(*~
	<docu>
		<summary>
			Parameter identifiers of the "Read parameters" command (manual pp. 43-46). Every value is exchanged as LONG x1000; times in seconds, levels in the instrument units, selections as code x1000.
		</summary>
	</docu>
~*)
{attribute 'qualified_only'}
{attribute 'strict'}
TYPE eTcoAteqG6_ParameterId_v_3_5_x :
(
	None := 0,
	FillTime := 1,
	StabTime := 2,
	TestTime := 3,
	PreFillTime := 6,
	DumpTime := 9,
	CouplingTimeA := 10,
	CouplingTimeB := 11,
	PartVolume := 20,
	TestType := 21,
	InterCycleTime := 29,
	ResultHoldTime := 48,
	MinFill := 50,
	MaxFill := 51,
	PressureUnit := 53,
	TestFail := 60,
	TestRework := 61,
	RefFail := 62,
	RefRework := 63,
	SetFill := 66,
	DiffAutoResetTime := 80,
	FillMode := 103,
	ExternalDumpType := 110,
	Input7Function := 112,
	Language := 123,
	MaxPreFill := 126,
	FlowUnit := 127,
	CalibrationLeakRate := 128,
	Filter := 148,
	UnitType := 149,
	BarGraphMaxReject := 158,
	VolumeUnit := 161,
	NextProgram := 164,
	PiezoAutoZeroCycles := 165,
	PiezoAutoZeroMinutes := 166,
	DelayExt1 := 249,
	DelayExt2 := 250,
	DelayExt3 := 251,
	DelayExt4 := 252,
	DelayExt5 := 253,
	DelayExt6 := 254,
	DelayInt2 := 255,
	DelayInt1 := 256,
	DelayAux1 := 257,
	DelayAux2 := 258,
	DelayAux3 := 259,
	DelayAux4 := 260,
	TimeExt1 := 261,
	TimeExt2 := 262,
	TimeExt3 := 263,
	TimeExt4 := 264,
	TimeExt5 := 265,
	TimeExt6 := 266,
	TimeInt2 := 267,
	TimeInt1 := 268,
	TimeAux1 := 269,
	TimeAux2 := 270,
	TimeAux3 := 271,
	TimeAux4 := 272,
	PressureFilter := 274,
	CapillaryRange := 281,
	BarCodeFirstChar := 287,
	BarCodeCharCount := 288,
	BarCodeProgram := 289,
	GeneralPressureUnit := 353,
	LinePressureMin := 354,
	DisplayMode := 364,
	Input8Function := 375,
	Input9Function := 376,
	UsbMode := 379,
	SaveOn := 412,
	AccessMode := 413,
	Year := 414,
	Month := 415,
	Day := 416,
	Hour := 417,
	Minute := 418,
	Second := 419,
	LearningCycles := 459,
	LearningInterCycleTime := 460,
	LearningMaxOffset := 461,
	LearningFlowMaster := 462,
	LearningPressureMaster := 463,
	LearningMinVolume := 464,
	LearningMaxVolume := 465,
	LearningOffset := 486
) UINT;
END_TYPE

(* stored: Version 1.1.0.1, ProductVersion 3.1.4024.12
   DUT eTcoAteqG6_ParameterId_v_3_5_x: Id {1d6f2124-6f40-4e6a-8469-e1ed0372d710} *)
